Fanuc KAREL source: kt00340.KL

-- PROVISIONAL review KL for V940-1; original PC SHA256 50bd832aa492dbf7059d595167273f99c585f04cefca8034a2f8d67992262d33
-- Incomplete behavior may be omitted. Consult companion uncertainty JSON. Do not deploy.
PROGRAM KT00340
%NOLOCKGROUP
VAR
  R2 : REAL
  OUT : BOOLEAN
-- UNRESOLVED_DECL Y1 type=002018
BEGIN
  -- V9_ZERO_TABLE_METADATA_HINT layout=0001; no indexed target words; source/name/runtime held
  -- UNRESOLVED_PC offsets 5-19; opcodes 2E,22,9D,33,B2
  -- UNRESOLVED_PC offsets 24-35; opcodes 2E,23
  -- UNRESOLVED_PC offsets 40-65; opcodes 22,9D,33,B1,21,29,64,29,6F,23
  -- UNRESOLVED_PC offsets 70-74; opcodes 7F
END KT00340
